(* IEC 61131-3 sources: plc-st-coding-agent/progress/evidence/f14_admission_preflight_20261111/native_artifacts/public-easy-05, 1 file *)

(* ---- candidate.st ---- *)
FUNCTION_BLOCK FB_WeldGapAlarm
VAR_INPUT
    Gap_Exceeded : BOOL;
    Weld_E_Stop_NC : BOOL;
    DebounceTime : TIME;
END_VAR
VAR_OUTPUT
    Operator_Alert : BOOL;
    Weld_Soft_Start_Active : BOOL;
END_VAR
VAR
    startupDelay : TON;
    gapDelay : TON;
END_VAR
startupDelay(IN := TRUE, PT := T#5s);
Weld_Soft_Start_Active := NOT startupDelay.Q;
gapDelay(IN := startupDelay.Q AND Weld_E_Stop_NC AND Gap_Exceeded, PT := DebounceTime);
Operator_Alert := gapDelay.Q;
END_FUNCTION_BLOCK
